TYPE ST_CamRecipe :
STRUCT
    lrObjectPitch : LREAL := 500.0;
    lrConveyorVelocity : LREAL := 100.0;
    lrCutVelocity : LREAL := 50.0;
    lrObjectEdgeLength : LREAL := 25.0;
    lrFirstEdgeStart : LREAL := 100.0;
    lrSecondEdgeStart : LREAL := 300.0;
    lrBlendMasterDistance : LREAL := 20.0;
    lrReturnEndPhase : LREAL := 480.0;
    lrMasterAcceleration : LREAL := 500.0;
    lrMasterDeceleration : LREAL := 500.0;
    lrMasterJerk : LREAL := 5000.0;
    lrMaxSlaveVelocity : LREAL := 600.0;
    lrMaxSlaveAcceleration : LREAL := 1600.0;
    lrMaxSlaveJerk : LREAL := 12000.0;
    lrRecoveryVelocity : LREAL := 100.0;
    lrRecoveryAcceleration : LREAL := 500.0;
    lrRecoveryDeceleration : LREAL := 500.0;
    lrRecoveryJerk : LREAL := 5000.0;
    lrPositionTolerance : LREAL := 0.1;
END_STRUCT
END_TYPE

(* stored: Version 1.1.0.1, ProductVersion 3.1.4024.16
   DUT ST_CamRecipe: Id {508fe896-e49a-47db-8cdd-6ac739ff50a2} *)
